// Integer field value of a typed publisher (PublishINT), BROTLib#4: the number with the trailing 'i'.
FUNCTION F_InfluxIntValue : STRING(255)
VAR_INPUT
	nValue		: LINT;
END_VAR

F_InfluxIntValue := CONCAT(LINT_TO_STRING(nValue), 'i');

END_FUNCTION

(* stored: Version 1.1.0.1, ProductVersion 3.1.4024.15
   POU F_InfluxIntValue: Id {132f3d79-4bf9-4f3d-bcf1-30bda9c04205}, SpecialFunc None *)
